(* IEC 61131-3 sources: plcassist-cli/packages/volt-lsp-iec/test-corpus/pro2193/Device/Plc Logic/Application/99 Library/Function Blocks/Actuators/Stacklights, Buttons, 9 files *)

(* ---- LedFB.fb ---- *)
// Control a colored led on a stacklight, or illuminated push-button
{attribute 'symbol' := 'none'}
FUNCTION_BLOCK PUBLIC LedFB
IMPLEMENTS IActuator, ILed
VAR
	Output			: ActuatorFB;
	FrequencySelect	: BOOL;
	xOverride		: BOOL;
	state			: enumLedState;
END_VAR

CASE state OF
	enumLedState.Off, enumLedState.ForcedOff:
		Output.Reset();

	enumLedState.Solid, enumLedState.ForcedOn:
		Output.Set();

	enumLedState.Flashing:
		IF NOT FrequencySelect THEN
			Output.SetOrReset(GlobalVars.BlinkerNormal);
		ELSE
			Output.SetOrReset(GlobalVars.BlinkerFast);
		END_IF

END_CASE

IF xOverride THEN
	Output.Set();
	xOverride := FALSE;
END_IF

// Instantiate the output
Output();

END_FUNCTION_BLOCK

// Start flashing the led
METHOD PUBLIC Flash
IF state <> enumLedState.ForcedOn AND state <> enumLedState.ForcedOff THEN
	state := enumLedState.Flashing;
END_IF
END_METHOD

// Force turn the led off
METHOD PUBLIC LedTestOff
state := enumLedState.ForcedOff;
END_METHOD

// Force turn the led on
METHOD PUBLIC LedTestOn
state := enumLedState.ForcedOn;
END_METHOD

// Stop forcing the led state
METHOD PUBLIC LedTestStop
state := enumLedState.Off;
END_METHOD

// Maps the actuator to the physical output
METHOD PUBLIC Map : BOOL
Map := Output.Map();
END_METHOD

// Turn the led off
METHOD PUBLIC Off
IF state <> enumLedState.ForcedOn AND state <> enumLedState.ForcedOff THEN
	state := enumLedState.Off;
END_IF
END_METHOD

// When button is pressed, set the led output without changing the state
METHOD PROTECTED Override
THIS^.xOverride := TRUE;
END_METHOD

// Reset the output (=False)
{attribute 'hide'}
METHOD Reset
Off();
END_METHOD

// Set the output (=True)
{attribute 'hide'}
METHOD Set : BOOL
Solid();
END_METHOD

METHOD PUBLIC SetFlashingFrequency
VAR_INPUT
	Value		: BOOL;		// Call with False to use (default) 0.5 sec. blinker. Call with True to use fast 0.2 sec. blinker.
END_VAR
FrequencySelect		:= Value;
END_METHOD

// Set the output True or False
METHOD SetOrReset
VAR_INPUT
	xValue	: BOOL;
END_VAR
IF xValue THEN
	state := enumLedState.Solid;
ELSE
	state := enumLedState.Off;
END_IF
END_METHOD

// Turn the led on
METHOD PUBLIC Solid
IF state <> enumLedState.ForcedOn AND state <> enumLedState.ForcedOff THEN
	state := enumLedState.Solid;
END_IF
END_METHOD

(* ---- PushButtonFunctionKeyFB.fb ---- *)
// Push button that is a function key (F1 or F2). Button sends extended state info to attached observers
FUNCTION_BLOCK PUBLIC PushButtonFunctionKeyFB
EXTENDS PushButtonLedFB
IMPLEMENTS IActuator, ISubject
VAR_INPUT
	buttonType				: enumHWButtons;	// The type of button will be supplied to attached observers
END_VAR
VAR
	Subject					: SubjectFunctionKeyFB;
	FunctionKeyState		:	// Keep internal state of function key
		(
			Released			:= 0,
			Tapped				:= 1,	// In state for as long as button is pressed, or until switched to Held
			AwaitingDoubleTap	:= 2,	// In state for max 1 sec.
			DoubleTapped		:= 3,	// In state for as long as button is pressed, or until switched to DoubleTapHeld
			Held				:= 4,
			DoubleTapHeld		:= 5,
		);
	HeldTrigger				: RisingTriggerFB;
	HeldTimer				: BTON;
	AwaitTapTimer			: BTON;
END_VAR
VAR CONSTANT
	HeldTimeout				: REAL := 0.5;		// Max 'Tap' duration. Switch to 'Held' state after this timeout
	AwaitTapTimeout			: REAL := 0.5;		// When released, await a double tap for this time.
END_VAR

// Implicit Enumeration: The implicit enumeration allows for an easy way to declare a new enumeration variable which is valid only within the local POU.
// https://content.helpme-codesys.com/en/CODESYS%20Development%20System/_cds_datatype_implicit_enumeration-1853150.html

SUPER^();

IF HeldTrigger.Rising(CLK := HeldTimer.Set(buttonInput, HeldTimeout)) THEN
	HandleHeld();
END_IF

IF AwaitTapTimer.Set(FunctionKeyState = AwaitingDoubleTap, AwaitTapTimeout) THEN
	FunctionKeyState := Released;
END_IF

END_FUNCTION_BLOCK

// Attach (subscribe) an observer to this subject. The observer will receive state from the subject.
METHOD PUBLIC Attach : BOOL
VAR_INPUT
	observer			: IObserver;
END_VAR
Attach := Subject.Attach(observer);
END_METHOD

// Detach (unsubscribe) an observer from this subject. The observer do longer receives updates.
METHOD PUBLIC Detach : BOOL
VAR_INPUT
	observer			: IObserver;
END_VAR
Detach := Subject.Detach(observer);
END_METHOD

METHOD PROTECTED HandleHeld
IF FunctionKeyState = Tapped THEN
	FunctionKeyState := Held;

	Subject.ButtonType	:= buttonType;
	Subject.ExtState	:= enumFunctionKeyPayload.Held;
	Subject.Notify();

ELSIF FunctionKeyState = DoubleTapped THEN
	FunctionKeyState := DoubleTapHeld;

	Subject.ButtonType	:= buttonType;
	Subject.ExtState	:= enumFunctionKeyPayload.DoubleTapHeld;
	Subject.Notify();

END_IF
END_METHOD

METHOD PROTECTED HandlePushed
SUPER^.HandlePushed();

IF FunctionKeyState = Released THEN
	FunctionKeyState := Tapped;
ELSIF FunctionKeyState = AwaitingDoubleTap THEN
	FunctionKeyState := DoubleTapped;
END_IF

Subject.ButtonType	:= buttonType;
Subject.ButtonState	:= TRUE;
Subject.ExtState	:= enumFunctionKeyPayload.Tapped;
Subject.Notify();
END_METHOD

METHOD PROTECTED HandleReleased
SUPER^.HandleReleased();

IF FunctionKeyState = Tapped THEN
	FunctionKeyState := AwaitingDoubleTap;
ELSIF FunctionKeyState = DoubleTapped THEN
	FunctionKeyState := Released;
ELSIF FunctionKeyState = Held OR FunctionKeyState = DoubleTapHeld THEN
	FunctionKeyState := Released;
END_IF

Subject.ButtonType	:= buttonType;
Subject.ButtonState	:= FALSE;
Subject.ExtState	:= enumFunctionKeyPayload.Released;
Subject.Notify();
END_METHOD

// The actual number of observers that are receiving events
{attribute 'monitoring' := 'call'}
PROPERTY ObserverCount : UINT
GET
VAR
END_VAR
ObserverCount := Subject.ObserverCount;
END_GET
END_PROPERTY

(* ---- PushButtonFunctionKeyFromCodesysVisuFB.fb ---- *)
// Push button from CODESYS WebVisu
FUNCTION_BLOCK PUBLIC PushButtonFunctionKeyFromCodesysVisuFB
EXTENDS PushButtonLedFB
IMPLEMENTS IActuator, ISubject
VAR_INPUT
	buttonType				: enumHWButtons;	// The type of button will be supplied to attached observers
END_VAR
VAR
	Subject					: SubjectFunctionKeyFromCodesysVisuFB;
	FunctionKeyState		:	// Keep internal state of function key
		(
			Released			:= 0,
			Tapped				:= 1,	// In state for as long as button is pressed, or until switched to Held
			AwaitingDoubleTap	:= 2,	// In state for max 1 sec.
			DoubleTapped		:= 3,	// In state for as long as button is pressed, or until switched to DoubleTapHeld
			Held				:= 4,
			DoubleTapHeld		:= 5,
		);
	HeldTrigger				: RisingTriggerFB;
	HeldTimer				: BTON;
	AwaitTapTimer			: BTON;
END_VAR
VAR CONSTANT
	HeldTimeout				: REAL := 0.5;		// Max 'Tap' duration. Switch to 'Held' state after this timeout
	AwaitTapTimeout			: REAL := 0.5;		// When released, await a double tap for this time.
END_VAR

// Implicit Enumeration: The implicit enumeration allows for an easy way to declare a new enumeration variable which is valid only within the local POU.
// https://content.helpme-codesys.com/en/CODESYS%20Development%20System/_cds_datatype_implicit_enumeration-1853150.html

SUPER^();

IF HeldTrigger.Rising(CLK := HeldTimer.Set(buttonInput, HeldTimeout)) THEN
	HandleHeld();
END_IF

IF AwaitTapTimer.Set(FunctionKeyState = AwaitingDoubleTap, AwaitTapTimeout) THEN
	FunctionKeyState := Released;
END_IF

END_FUNCTION_BLOCK

// Attach (subscribe) an observer to this subject. The observer will receive state from the subject.
METHOD PUBLIC Attach : BOOL
VAR_INPUT
	observer			: IObserver;
END_VAR
Attach := Subject.Attach(observer);
END_METHOD

// Detach (unsubscribe) an observer from this subject. The observer do longer receives updates.
METHOD PUBLIC Detach : BOOL
VAR_INPUT
	observer			: IObserver;
END_VAR
Detach := Subject.Detach(observer);
END_METHOD

METHOD PROTECTED HandleHeld
IF FunctionKeyState = Tapped THEN
	FunctionKeyState := Held;

	Subject.ButtonType	:= buttonType;
	Subject.ExtState	:= enumFunctionKeyPayload.Held;
	Subject.Notify();

ELSIF FunctionKeyState = DoubleTapped THEN
	FunctionKeyState := DoubleTapHeld;

	Subject.ButtonType	:= buttonType;
	Subject.ExtState	:= enumFunctionKeyPayload.DoubleTapHeld;
	Subject.Notify();

END_IF
END_METHOD

METHOD PROTECTED HandlePushed
SUPER^.HandlePushed();

IF FunctionKeyState = Released THEN
	FunctionKeyState := Tapped;
ELSIF FunctionKeyState = AwaitingDoubleTap THEN
	FunctionKeyState := DoubleTapped;
END_IF

Subject.ButtonType	:= buttonType;
//Subject.ButtonState	:= TRUE;
Subject.ExtState	:= enumFunctionKeyPayload.Tapped;
Subject.Notify();
END_METHOD

METHOD PROTECTED HandleReleased
SUPER^.HandleReleased();

IF FunctionKeyState = Tapped THEN
	FunctionKeyState := AwaitingDoubleTap;
ELSIF FunctionKeyState = DoubleTapped THEN
	FunctionKeyState := Released;
ELSIF FunctionKeyState = Held OR FunctionKeyState = DoubleTapHeld THEN
	FunctionKeyState := Released;
END_IF

Subject.ButtonType	:= buttonType;
//Subject.ButtonState	:= FALSE;
Subject.ExtState	:= enumFunctionKeyPayload.Released;
Subject.Notify();
END_METHOD

// The actual number of observers that are receiving events
{attribute 'monitoring' := 'call'}
PROPERTY ObserverCount : UINT
GET
VAR
END_VAR
ObserverCount := Subject.ObserverCount;
END_GET
END_PROPERTY

(* ---- PushButtonLedFB.fb ---- *)
// Control an illuminated push-button
{attribute 'symbol' := 'none'}
FUNCTION_BLOCK PUBLIC PushButtonLedFB
EXTENDS LedFB
IMPLEMENTS IActuator
VAR_INPUT
	buttonInput				: BOOL;			// Connect to hardware
END_VAR
VAR
	{attribute 'hide'}
	Trig_Pushed				: TriggerFB;
END_VAR

CallTrigger();

IF ButtonPushed THEN
	HandlePushed();
END_IF

IF buttonInput THEN	// Illuminate button while pressed down
	Override();
END_IF

IF ButtonReleased THEN
	HandleReleased();
END_IF

SUPER^();

END_FUNCTION_BLOCK

METHOD PROTECTED CallTrigger
Trig_Pushed.Call(CLK := buttonInput);
END_METHOD

METHOD PROTECTED HandlePushed
//savedState := State;
//Solid();
END_METHOD

METHOD PROTECTED HandleReleased
//State := savedState;
END_METHOD

// Give a signal on rising edge when the button is pushed.
PROPERTY PUBLIC ButtonPushed : BOOL
GET
VAR
END_VAR
ButtonPushed := Trig_Pushed.Q_Rising;
END_GET
END_PROPERTY

// Give a signal on faling edge when the button is released.
PROPERTY PUBLIC ButtonReleased : BOOL
GET
VAR
END_VAR
ButtonReleased := Trig_Pushed.Q_Falling;
END_GET
END_PROPERTY

(* ---- PushButtonLedWithHmiFB.fb ---- *)
// Control an illuminated push-button, also handle input from the visualisation. Set the color of the button.
// Remember to declare this FB with: '{attribute 'symbol' := 'readwrite'}'
{attribute 'symbol' := 'none'}
FUNCTION_BLOCK PUBLIC PushButtonLedWithHmiFB
EXTENDS PushButtonLedFB
IMPLEMENTS IActuator
VAR
	{attribute 'symbol' := 'readwrite'}	button					: BOOL;				// Button is pushed down (from HMI)
	{attribute 'symbol' := 'read'}		feedback				: enumColorList;	// Current color of button

	colorOn			: enumColorList		:= enumColorList.Lime;
	colorOff		: enumColorList		:= enumColorList.Silver;
	colorPushed		: enumColorList		:= enumColorList.Black;
END_VAR

// Illuminate button while pressed down
IF button THEN
	Override();
END_IF

CASE state OF
	enumLedState.Off, enumLedState.ForcedOff:
		feedback		:= colorOff;

	enumLedState.Solid, enumLedState.ForcedOn:
		feedback		:= colorOn;

	enumLedState.Flashing:
		IF NOT FrequencySelect THEN
			feedback	:= SEL(GlobalVars.BlinkerNormal, colorOff, colorOn);
		ELSE
			feedback	:= SEL(GlobalVars.BlinkerFast, colorOff, colorOn);
		END_IF

END_CASE

IF xOverride THEN
	feedback := colorPushed;
END_IF

SUPER^();

END_FUNCTION_BLOCK

METHOD PROTECTED CallTrigger
Trig_Pushed.Call(CLK := buttonInput OR button);
END_METHOD

// Set the colors for the button
METHOD PUBLIC SetColors
VAR_INPUT
	colorOn			: enumColorList		:= enumColorList.Lime;
	colorOff		: enumColorList		:= enumColorList.Silver;
	colorPushed		: enumColorList		:= enumColorList.Black;
END_VAR
THIS^.colorOn			:= colorOn;
THIS^.colorOff			:= colorOff;
THIS^.colorPushed		:= colorPushed;
END_METHOD

(* ---- PushButtonWithObserverFB.fb ---- *)
// Push button that is any of the buttons defined in enumHWButtons. Button sends state to attached observers
FUNCTION_BLOCK PUBLIC PushButtonWithObserverFB
EXTENDS PushButtonLedFB
IMPLEMENTS IActuator, ISubject
VAR_INPUT
	buttonType				: enumHWButtons;	// The type of button will be supplied to attached observers
END_VAR
VAR
	Subject					: SubjectHWButtonFB;
END_VAR

SUPER^();

END_FUNCTION_BLOCK

// Attach (subscribe) an observer to this subject. The observer will receive state from the subject.
METHOD PUBLIC Attach : BOOL
VAR_INPUT
	observer			: IObserver;
END_VAR
Attach := Subject.Attach(observer);
END_METHOD

// Detach (unsubscribe) an observer from this subject. The observer do longer receives updates.
METHOD PUBLIC Detach : BOOL
VAR_INPUT
	observer			: IObserver;
END_VAR
Detach := Subject.Detach(observer);
END_METHOD

METHOD PROTECTED HandlePushed
SUPER^.HandlePushed();

Subject.ButtonType	:= buttonType;
Subject.ButtonState	:= TRUE;
Subject.Notify();
END_METHOD

METHOD PROTECTED HandleReleased
SUPER^.HandleReleased();

Subject.ButtonType	:= buttonType;
Subject.ButtonState	:= FALSE;
Subject.Notify();
END_METHOD

// The actual number of observers that are receiving events
{attribute 'monitoring' := 'call'}
PROPERTY ObserverCount : UINT
GET
VAR
END_VAR
ObserverCount := Subject.ObserverCount;
END_GET
END_PROPERTY

(* ---- StacklightFB.fb ---- *)
// Control a stacklight with several colored lamps, and a buzzer
FUNCTION_BLOCK PUBLIC StacklightFB
IMPLEMENTS IActuator
VAR_INPUT
	Green			: LedFB;
	Amber			: LedFB;
	Red				: LedFB;
END_VAR
VAR
END_VAR

// Instantiate the outputs
Green();
Amber();
Red();

END_FUNCTION_BLOCK

// Maps the actuator to the physical output
{attribute 'hide'}
METHOD PUBLIC Map : BOOL
// no implementation
END_METHOD

// Reset all outputs on the stacklight
METHOD Reset
Green.Off();
Amber.Off();
Red.Off();
END_METHOD

// Set the output (=True)
{attribute 'hide'}
METHOD Set : BOOL
// no implementation
END_METHOD

// Set the output True or False
{attribute 'hide'}
METHOD SetOrReset
VAR_INPUT
	xValue	: BOOL;
END_VAR
// no implementation
END_METHOD

(* ---- StacklightWithBlueFB.fb ---- *)
// Control a stacklight with several colored lamps, and a buzzer
FUNCTION_BLOCK PUBLIC StacklightWithBlueFB
EXTENDS StacklightFB
IMPLEMENTS IActuator
VAR_INPUT
	Blue			: LedFB;
END_VAR

// Instantiate the outputs
SUPER^();
Blue();

END_FUNCTION_BLOCK

// Reset all outputs on the stacklight
METHOD Reset
SUPER^.Reset();
Blue.Off();
END_METHOD

(* ---- StacklightWithHornFB.fb ---- *)
// Control a stacklight with several colored lamps, and a buzzer
FUNCTION_BLOCK PUBLIC StacklightWithHornFB
EXTENDS StacklightFB
IMPLEMENTS IActuator
VAR_INPUT
	Horn			: LedFB;
END_VAR

// Instantiate the outputs
SUPER^();
Horn();

END_FUNCTION_BLOCK

// Reset all outputs on the stacklight
METHOD Reset
SUPER^.Reset();
Horn.Off();
END_METHOD
